Fanuc KAREL source: KT00481.KL

PROGRAM KT00481
%NOLOCKGROUP
VAR
  P1: POSITION
  P2: XYZWPR
  OUT: XYZWPREXT
BEGIN
    P2.Y = 2.0
  OUT = P1 : P2
END KT00481
